FUNCTION_BLOCK FB_YASKAWA_Controller
(*

The function block used to control axis.

Constructor: 		Patryk Panylo
Company:		E. Riexinger GmbH
Date:			20.06.2018
Version:			1.00

Date:			Revision:		Who:				Comment
dd.mm.yyyy		x.xx			Initials			comment

*)
VAR_INPUT
	(* Input variables / Eingang Variablen *)
	bEnable						:BOOL;						(* Signal FB enable *)
	etMachineMode				:ET_MachineMode;			(* Machine mode *)
	etMachineState				:ET_MachineState;			(* Machine state *)
	bDrivesOn					:BOOL;						(* Enable the drives *)
	bMoveOn					:BOOL;						(* Enable the move enable *)
	bReset						:BOOL;						(* Signal reset *)
	bExeReset					:BOOL;						(* Execute auto reset *)
	lrOverride					:LREAL;						(* Override 100% percent *)
END_VAR
VAR_OUTPUT
	(* Output variables / Ausgang Variablen *)
	bStatus						:BOOL;						(* Feedback *)
	bStatusDelay					:BOOL;						(* Feedback delay *)
	bReseted					:BOOL;						(* Reset completed *)
	bError						:BOOL;						(* Controller error *)
	udnErrorNo					:UDINT;						(* Error number *)
	bInHome						:BOOL;						(* In home *)
	bNotMoving					:BOOL;						(* Status of moving *)
	bNotInCrashAreaMachine		:BOOL;						(* Status not in crash area *)
END_VAR
VAR_IN_OUT
	(* Input Output variables / Ausgang Variablen *)
	Yaskawa					:ST_YASKAWA_REF;				(* The YASKAWA_REF data type  is an interface between the PLC and the YASKAWA and contains axis information *)
END_VAR
VAR
	(* Enummerations *)

	(* Variables *)
	tStatusDelay					:TIME := t#1s;					(* Status delay time *)

	bFirstTime					:BOOL;

	(* References *)

	(* Interfaces *)

	(* Instances *)
	fbPower						:FB_YASKAWA_Power;		(* The function block is used to enable for an axis *)
	tonStatusDelay				:TON;						(* Delay controller enabled status *)
	fbReset						:FB_YASKAWA_Reset;			(* An axis reset is carried out with the function block *)

END_VAR


IF NOT bEnable							(* Signal FB enable *)
THEN
	bStatus := FALSE;						(* Feedback *)
	bStatusDelay := FALSE;				(* Feedback *)
	bError := FALSE;						(* Controller error *)
	udnErrorNo := 0;						(* Error number *)

	bFirstTime := FALSE;
	RETURN;
END_IF

IF NOT bFirstTime
THEN

	bFirstTime := TRUE;
END_IF;

A_Power();
A_Reset();
A_Error();

(* In home *)
bInHome := Yaskawa.stYaskawaToPlc.bInHome;

(* Status not moving *)
bNotMoving := Yaskawa.stYaskawaToPlc.bNotMoving;

(* Status not in crash area *)
bNotInCrashAreaMachine := Yaskawa.stYaskawaToPlc.bNotInCrashAreaMachine;

ACTION A_Error:

bError := fbReset.bError
	         OR fbPower.bError;
END_ACTION

ACTION A_Power:

fbPower(
	bEnable := TRUE,
	bAutoHand := etMachineMode = ET_MachineMode_eHome
			         OR etMachineMode = ET_MachineMode_eStepping
			         OR etMachineMode = ET_MachineMode_eAutomatic,
	bDrivesOn :=  bDrivesOn,
	bMoveOn := bMoveOn,
	lrOverride := lrOverride,
	Yaskawa := Yaskawa
 );

tonStatusDelay(
	IN := fbPower.bStatus,
	PT := SEL(etMachineMode = ET_MachineMode_eManual, tStatusDelay, t#0ms),
	Q => bStatusDelay
);
END_ACTION

ACTION A_Reset:

fbReset(
	bExecute := bReset
	            	     XOR bExeReset,
	Yaskawa := Yaskawa,
	bDone => bReseted
);
END_ACTION

END_FUNCTION_BLOCK

(* stored: Version 1.1.0.1, ProductVersion 3.1.4024.15
   POU FB_YASKAWA_Controller: Id {ea52ded9-74c3-4ead-be54-16fd37ad7735}, SpecialFunc None
   Action A_Error: Id {2788d67a-913c-4651-98e7-7a554302a478}
   Action A_Power: Id {9bb3910a-abbb-4409-865a-f134bbc02d84}
   Action A_Reset: Id {bc3ab0da-783f-47ea-93c6-583262356a74} *)
